(* IEC 61131-3 sources: STruCpp/tests/st-validation/functions, 8 files *)

(* ---- basic_function.st ---- *)
FUNCTION AddInts : INT
  VAR_INPUT a : INT; b : INT; END_VAR
  AddInts := a + b;
END_FUNCTION

FUNCTION IsPositive : BOOL
  VAR_INPUT val : INT; END_VAR
  IsPositive := val > 0;
END_FUNCTION

FUNCTION MaxInt : INT
  VAR_INPUT a : INT; b : INT; END_VAR
  IF a > b THEN
    MaxInt := a;
  ELSE
    MaxInt := b;
  END_IF;
END_FUNCTION

(* ---- function_calls.st ---- *)
FUNCTION Double : INT
  VAR_INPUT x : INT; END_VAR
  Double := x * 2;
END_FUNCTION

FUNCTION Triple : INT
  VAR_INPUT x : INT; END_VAR
  Triple := x * 3;
END_FUNCTION

FUNCTION_BLOCK Calculator
  VAR_INPUT base : INT; END_VAR
  VAR_OUTPUT doubled : INT; tripled : INT; END_VAR
  doubled := Double(x := base);
  tripled := Triple(x := base);
END_FUNCTION_BLOCK

(* ---- bitwise_mixed.st ---- *)
PROGRAM BitwiseMixed
  VAR
    and_dw : DWORD;
    or_dw : DWORD;
    xor_dw : DWORD;
    and3_dw : DWORD;
    mixed_or_dw : DWORD;
  END_VAR

  and_dw := AND(DWORD#16#000000FF, WORD#16#00FF);
  or_dw := OR(DWORD#16#000000FF, WORD#16#00FF);
  xor_dw := XOR(DWORD#16#0000000F, WORD#16#00F0);
  and3_dw := AND(DWORD#16#00FF, WORD#16#000F, BYTE#16#03);
  mixed_or_dw := OR(WORD#16#00FF, DWORD#16#FF00);
END_PROGRAM

(* ---- std_functions.st ---- *)
PROGRAM StdFunctionsTest
  VAR
    abs_result : INT;
    min_result : INT;
    max_result : INT;
    a : INT;
    b : INT;
    c : INT;
    flag_a : BOOL := TRUE;
    flag_b : BOOL := FALSE;
    flag_c : BOOL := TRUE;
    and_result : BOOL;
    and3_result : BOOL;
    or_result : BOOL;
    xor_result : BOOL;
    not_result : BOOL;
    mod_result : INT;
    infix_and : BOOL;
    infix_or : BOOL;
    infix_not : BOOL;
    infix_mod : INT;
  END_VAR

  a := -42;
  b := 10;
  c := 3;
  abs_result := ABS(a);
  min_result := MIN(b, c);
  max_result := MAX(b, c);

  (* Operator keywords used as function calls — FBD-style *)
  and_result := AND(flag_a, flag_b);
  and3_result := AND(flag_a, flag_b, flag_c);
  or_result := OR(flag_a, flag_b);
  xor_result := XOR(flag_a, flag_b);
  not_result := NOT(flag_a);
  mod_result := MOD(b, c);

  (* Infix operators must still work alongside function-call form *)
  infix_and := flag_a AND flag_b;
  infix_or := flag_a OR flag_b;
  infix_not := NOT flag_a;
  infix_mod := b MOD c;
END_PROGRAM

(* ---- test_basic_function.st ---- *)
TEST 'Add two positive integers'
  VAR result : INT; END_VAR
  result := AddInts(a := 3, b := 7);
  ASSERT_EQ(result, 10);
END_TEST

TEST 'Add with negative'
  VAR result : INT; END_VAR
  result := AddInts(a := -5, b := 3);
  ASSERT_EQ(result, -2);
END_TEST

TEST 'Add zeros'
  VAR result : INT; END_VAR
  result := AddInts(a := 0, b := 0);
  ASSERT_EQ(result, 0);
END_TEST

TEST 'IsPositive true'
  VAR result : BOOL; END_VAR
  result := IsPositive(val := 5);
  ASSERT_TRUE(result);
END_TEST

TEST 'IsPositive false for zero'
  VAR result : BOOL; END_VAR
  result := IsPositive(val := 0);
  ASSERT_FALSE(result);
END_TEST

TEST 'Max returns larger value'
  VAR result : INT; END_VAR
  result := MaxInt(a := 10, b := 20);
  ASSERT_EQ(result, 20);
END_TEST

TEST 'Max with equal values'
  VAR result : INT; END_VAR
  result := MaxInt(a := 5, b := 5);
  ASSERT_EQ(result, 5);
END_TEST

(* ---- test_bitwise_mixed.st ---- *)
TEST 'AND with mixed bit types'
  VAR uut : BitwiseMixed; END_VAR
  uut();
  ASSERT_EQ(uut.and_dw, 255);
END_TEST

TEST 'OR with mixed bit types'
  VAR uut : BitwiseMixed; END_VAR
  uut();
  ASSERT_EQ(uut.or_dw, 255);
END_TEST

TEST 'XOR with mixed bit types'
  VAR uut : BitwiseMixed; END_VAR
  uut();
  ASSERT_EQ(uut.xor_dw, 255);
END_TEST

TEST 'AND variadic with mixed bit types'
  VAR uut : BitwiseMixed; END_VAR
  uut();
  ASSERT_EQ(uut.and3_dw, 3);
END_TEST

TEST 'OR with smaller first operand'
  VAR uut : BitwiseMixed; END_VAR
  uut();
  ASSERT_EQ(uut.mixed_or_dw, 65535);
END_TEST

(* ---- test_function_calls.st ---- *)
TEST 'Direct function call'
  VAR result : INT; END_VAR
  result := Double(x := 7);
  ASSERT_EQ(result, 14);
END_TEST

TEST 'Function called from FB'
  VAR calc : Calculator; END_VAR
  calc(base := 5);
  ASSERT_EQ(calc.doubled, 10);
  ASSERT_EQ(calc.tripled, 15);
END_TEST

TEST 'Nested function calls in expression'
  VAR result : INT; END_VAR
  result := Double(x := Triple(x := 2));
  ASSERT_EQ(result, 12);
END_TEST

(* ---- test_std_functions.st ---- *)
TEST 'ABS of negative'
  VAR uut : StdFunctionsTest; END_VAR
  uut();
  ASSERT_EQ(uut.abs_result, 42);
END_TEST

TEST 'MIN returns smaller'
  VAR uut : StdFunctionsTest; END_VAR
  uut();
  ASSERT_EQ(uut.min_result, 3);
END_TEST

TEST 'MAX returns larger'
  VAR uut : StdFunctionsTest; END_VAR
  uut();
  ASSERT_EQ(uut.max_result, 10);
END_TEST

TEST 'AND function call (2 args)'
  VAR uut : StdFunctionsTest; END_VAR
  uut();
  ASSERT_EQ(uut.and_result, FALSE);
END_TEST

TEST 'AND function call (3 args variadic)'
  VAR uut : StdFunctionsTest; END_VAR
  uut();
  ASSERT_EQ(uut.and3_result, FALSE);
END_TEST

TEST 'OR function call'
  VAR uut : StdFunctionsTest; END_VAR
  uut();
  ASSERT_EQ(uut.or_result, TRUE);
END_TEST

TEST 'XOR function call'
  VAR uut : StdFunctionsTest; END_VAR
  uut();
  ASSERT_EQ(uut.xor_result, TRUE);
END_TEST

TEST 'NOT function call'
  VAR uut : StdFunctionsTest; END_VAR
  uut();
  ASSERT_EQ(uut.not_result, FALSE);
END_TEST

TEST 'MOD function call'
  VAR uut : StdFunctionsTest; END_VAR
  uut();
  ASSERT_EQ(uut.mod_result, 1);
END_TEST

TEST 'infix AND matches function-call AND'
  VAR uut : StdFunctionsTest; END_VAR
  uut();
  ASSERT_EQ(uut.infix_and, uut.and_result);
END_TEST

TEST 'infix OR matches function-call OR'
  VAR uut : StdFunctionsTest; END_VAR
  uut();
  ASSERT_EQ(uut.infix_or, uut.or_result);
END_TEST

TEST 'infix NOT matches function-call NOT'
  VAR uut : StdFunctionsTest; END_VAR
  uut();
  ASSERT_EQ(uut.infix_not, uut.not_result);
END_TEST

TEST 'infix MOD matches function-call MOD'
  VAR uut : StdFunctionsTest; END_VAR
  uut();
  ASSERT_EQ(uut.infix_mod, uut.mod_result);
END_TEST
